// TIA Portal V20 export
// export: Created 2026-11-24T19:16:26.3193844Z, ExportSetting WithDefaults, DisplayName Totally Integrated Automation Portal, DisplayVersion V20 Update 7, DisplayName TIA Portal Openness, DisplayVersion V20 Update 7, DisplayName TIA Portal Version Control Interface, DisplayVersion V20 Update 7, DisplayName TIA Portal Test Suite Advanced, DisplayVersion V20, DisplayName SINAMICS Startdrive Advanced, DisplayVersion V20 SP1 Update 1, DisplayName SINAMICS Startdrive G110M, G120, G120C, G120D, G120P, G115D, DisplayVersion V20 SP1 Update 1, DisplayName SINAMICS Startdrive G130, G150, S120, S150, SINAMICS MV, G220, S200, S210, DisplayVersion V20 SP1 Update 1, DisplayName STEP 7 Professional, DisplayVersion V20 Update 7, DisplayName STEP 7 Safety, DisplayVersion V20 Update 2, DisplayName WinCC Basic/Comfort/Advanced, DisplayVersion V20 Update 7, DisplayName WinCC Unified, DisplayVersion V20 Update 7
FUNCTION_BLOCK "zzLadControl"   // FB5, LAD
{ S7_Optimized_Access := 'TRUE' }
VERSION : 0.1
// Inventory: Program control operations
// stored: AutoNumber true, IsIECCheckEnabled false, IsRetainMemResEnabled false, MemoryReserve 100, SetENOAutomatically false, UDAEnableTagReadback false
BEGIN

REGION Network 1: CoilRetValue
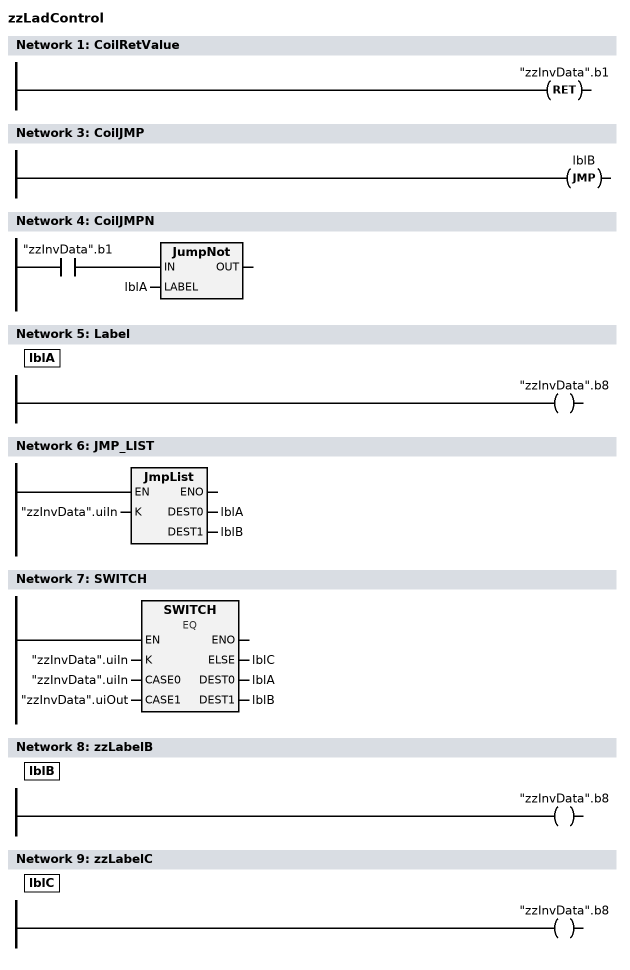
   ENO := "zzInvData".b1;
   RETURN;
END_REGION

REGION Network 2: Empty
END_REGION

REGION Network 3: CoilJMP
   RUNG wire#powerrail
      JumpCoil( lblB )
   END_RUNG
   // the same network as SCL:
   GOTO lblB;
END_REGION

REGION Network 4: CoilJMPN
   // no SCL statement known for JumpNot: written as a call
   JumpNot(in := "zzInvData".b1, label := lblA);
END_REGION

REGION Network 5: Label
   Label( lblA )
   RUNG wire#powerrail
      Coil( "zzInvData".b8 )
   END_RUNG
   // the same network as SCL:
   lblA:
   "zzInvData".b8 := TRUE;
END_REGION

REGION Network 6: JMP_LIST
   // no SCL statement known for JmpList: written as a call
   JmpList(k := "zzInvData".uiIn, dest0 => lblA, dest1 => lblB);
END_REGION

REGION Network 7: SWITCH
   // no SCL statement known for Switch: written as a call
   Switch(k := "zzInvData".uiIn,
          case0 := "zzInvData".uiIn,
          case1 := "zzInvData".uiOut,
          "else" => lblC,
          dest0 => lblA,
          dest1 => lblB);
END_REGION

REGION Network 8: zzLabelB
   Label( lblB )
   RUNG wire#powerrail
      Coil( "zzInvData".b8 )
   END_RUNG
   // the same network as SCL:
   lblB:
   "zzInvData".b8 := TRUE;
END_REGION

REGION Network 9: zzLabelC
   Label( lblC )
   RUNG wire#powerrail
      Coil( "zzInvData".b8 )
   END_RUNG
   // the same network as SCL:
   lblC:
   "zzInvData".b8 := TRUE;
END_REGION
END_FUNCTION_BLOCK
